(* IEC 61131-3 sources: stf-hw/stf-cad/line2/plc, 16 files *)

(* ---- DUT_PhysicalAI.st ---- *)
// timestamped I/O and the record every learned model is trained on
TYPE ST_TsInput : STRUCT bNewEdge : BOOL; nTimestamp : ULINT; END_STRUCT; END_TYPE     // EL1252 (DC ns)
TYPE ST_TsOutput : STRUCT bArm : BOOL; nFireAt : ULINT; END_STRUCT; END_TYPE          // EL2252 (DC ns)
// station states: named types (an enumeration declared inline in a VAR block is not portable)
TYPE T_ZoneArray : ARRAY[0..2] OF LREAL; END_TYPE   // per oven zone (one named type: FB_Band -> FB_Oven)
TYPE E_PickState : (WAIT, TRACK, GRIP, LIFT, PLACE, RELEASE, HOME); END_TYPE
TYPE E_AirlockOut : (IDLE, CARRY_OUT, INNER_CLOSE, OUTER_OPEN, SWAP, OUTER_CLOSE, INNER_OPEN, CARRY_IN); END_TYPE
// the stations (DT-4b)
TYPE ST_DeltaJob : STRUCT              // PLC -> a delta's motion program: a new nJob starts the job
    nJob : INT; nPuck : INT; nCol : INT; nLane : INT;   // C: the band row (fRowPos) + column -> puck; A/B: puck -> lane
    fRowPos : LREAL; fStart : LREAL;                    // band mm of the row's cut; master mm to start at
END_STRUCT; END_TYPE
TYPE ST_QcResult : STRUCT nSeq : INT; nPuck : INT; nVerdict : INT; END_STRUCT; END_TYPE   // edge PC: 1 pass, 2 reject
TYPE ST_Puck : STRUCT
    bFull : BOOL; bKicked : BOOL; bPending : BOOL;      // pending: a pick is decided, its grip not yet known
    nFlav : INT; nCol : INT; nVerdict : INT; fRowPos : LREAL;
END_STRUCT; END_TYPE
TYPE T_PuckArray : ARRAY[0..47] OF ST_Puck; END_TYPE
TYPE ST_Lane : STRUCT fBlock : LREAL; fPackAt : LREAL; nPackReq : INT; bCanPack : BOOL; END_STRUCT; END_TYPE   // s (master)
TYPE T_LaneArray : ARRAY[0..2] OF ST_Lane; END_TYPE
TYPE ST_PuckEvent : STRUCT
    nPuck : UINT; sNfc : STRING(16); nDcTime : ULINT; fMasterPos : LREAL;
    eStation : E_Station; aSignals : ARRAY[0..15] OF REAL; nImageId : UDINT; eOutcome : E_Outcome;
END_STRUCT; END_TYPE

(* ---- GVL_IO.st ---- *)
// GVL_IO - generated by plc_io.py from line_model: every signal, mapped in the I/O tree
{attribute 'qualified_only'}
VAR_GLOBAL
    axQ1                            : AXIS_REF;   // -KF20 ch1      M1_master_drive              stepper 17HS19-2004D-E1000+PG27
    encB1                    AT %I* : UDINT;   // -KF18 ch1      B1_master_encoder            master encoder, 1024 ppr RS422
    axQ41                           : AXIS_REF;   // -KF21 ch1      M_dep_rolls                  stepper 17HS19-2004D-E1000+PG27
    iolIOL1                  AT %I* : INT;   // -KF14 ch1      dep_hopper_level             ToF level (IO-Link)
    qQ2                      AT %Q* : BOOL;   // -KF5 ch7       top_cyl_weiss                valve coil (ISO6432-16x25)
    iQ2_S1                   AT %I* : BOOL;   // -KF1 ch1       top_cyl_weiss                reed switch retracted (ISO6432-16x25)
    iQ2_S2                   AT %I* : BOOL;   // -KF1 ch2       top_cyl_weiss                reed switch extended (ISO6432-16x25)
    qQ3                      AT %Q* : BOOL;   // -KF5 ch8       top_cyl_rot                  valve coil (ISO6432-16x25)
    iQ3_S1                   AT %I* : BOOL;   // -KF1 ch3       top_cyl_rot                  reed switch retracted (ISO6432-16x25)
    iQ3_S2                   AT %I* : BOOL;   // -KF1 ch4       top_cyl_rot                  reed switch extended (ISO6432-16x25)
    qQ4                      AT %Q* : BOOL;   // -KF5 ch9       top_cyl_blau                 valve coil (ISO6432-16x25)
    iQ4_S1                   AT %I* : BOOL;   // -KF1 ch5       top_cyl_blau                 reed switch retracted (ISO6432-16x25)
    iQ4_S2                   AT %I* : BOOL;   // -KF1 ch6       top_cyl_blau                 reed switch extended (ISO6432-16x25)
    iolIOL5                  AT %I* : INT;   // -KF14 ch2      top_level_weiss              ToF level (IO-Link)
    iolIOL6                  AT %I* : INT;   // -KF14 ch3      top_level_rot                ToF level (IO-Link)
    iolIOL7                  AT %I* : INT;   // -KF14 ch4      top_level_blau               ToF level (IO-Link)
    axQ40                           : AXIS_REF;   // -KF22 ch1      M_band                       stepper 17HS19-2004D-E1000+PG27
    qE1T1                    AT %Q* : BOOL;   // -KF5 ch12      oven_heater_E1T1             oven element SSR (500 W 230 V, L1)
    qE1T2                    AT %Q* : BOOL;   // -KF5 ch13      oven_heater_E1T2             oven element SSR (500 W 230 V, L2)
    qE1T3                    AT %Q* : BOOL;   // -KF5 ch14      oven_heater_E1T3             oven element SSR (500 W 230 V, L3)
    qE1B1                    AT %Q* : BOOL;   // -KF5 ch10      oven_heater_E1B1             oven element SSR (500 W 230 V, L1)
    qE1B2                    AT %Q* : BOOL;   // -KF5 ch11      oven_heater_E1B2             oven element SSR (500 W 230 V, L2)
    qQF1                     AT %Q* : BOOL;   // -KF6 ch7       oven_fan_1_motor             oven circulation fan 230 V 35 W (L2), coupling relay
    tcTC1                    AT %I* : INT;   // -KF12 ch1      oven_tc_1                    oven zone thermocouple K (duplex: this element -> PID)
    qE2T1                    AT %Q* : BOOL;   // -KF5 ch16      oven_heater_E2T1             oven element SSR (500 W 230 V, L3)
    qE2B1                    AT %Q* : BOOL;   // -KF5 ch15      oven_heater_E2B1             oven element SSR (350 W 230 V, L2)
    qQF2                     AT %Q* : BOOL;   // -KF6 ch8       oven_fan_2_motor             oven circulation fan 230 V 35 W (L3), coupling relay
    tcTC2                    AT %I* : INT;   // -KF12 ch2      oven_tc_2                    oven zone thermocouple K (duplex: this element -> PID)
    qE3T1                    AT %Q* : BOOL;   // -KF6 ch2       oven_heater_E3T1             oven element SSR (500 W 230 V, L1)
    qE3B1                    AT %Q* : BOOL;   // -KF6 ch1       oven_heater_E3B1             oven element SSR (350 W 230 V, L3)
    qQF3                     AT %Q* : BOOL;   // -KF6 ch9       oven_fan_3_motor             oven circulation fan 230 V 35 W (L2), coupling relay
    tcTC3                    AT %I* : INT;   // -KF12 ch3      oven_tc_3                    oven zone thermocouple K (duplex: this element -> PID)
    qQX1                     AT %Q* : BOOL;   // -KF6 ch10      oven_exhaust_fan             oven vapour exhaust fan 24 V EC
    aiIR1                    AT %I* : INT;   // -KF9 ch4       IR1_pyrometer                product temperature 0..10 V
    qQC1                     AT %Q* : BOOL;   // -KF6 ch3       cool_fan_1                   band cooling fan 24 V
    qQC2                     AT %Q* : BOOL;   // -KF6 ch4       cool_fan_2                   band cooling fan 24 V
    qQC3                     AT %Q* : BOOL;   // -KF6 ch5       cool_exfan_1                 band cooling fan 24 V
    qQC4                     AT %Q* : BOOL;   // -KF6 ch6       cool_exfan_2                 band cooling fan 24 V
    axdelta_C_M60                   : AXIS_REF;   // -KF25 ch1      delta_C_motor_60             stepper 17HS19-2004D-E1000+SWG17-30
    axdelta_C_M180                  : AXIS_REF;   // -KF23 ch1      delta_C_motor_180            stepper 17HS19-2004D-E1000+SWG17-30
    axdelta_C_M300                  : AXIS_REF;   // -KF24 ch1      delta_C_motor_300            stepper 17HS19-2004D-E1000+SWG17-30
    qdelta_C_VAC             AT %Q* : BOOL;   // -KF6 ch11      delta_C_cup_a                vacuum ejector valve
    ioldelta_C_VAC_P         AT %I* : INT;   // -KF15 ch2      delta_C_cup_a                vacuum level (analogue grip quality)
    iI1                      AT %I* : BOOL;   // -KF1 ch13      I1_full_check                puck already full (recirculating) -> delta C does NOT place
    iolNFC_W                 AT %I* : ARRAY[0..31] OF BYTE;   // -KF15 ch1      nfc_writer                   RFID/NFC head (IO-Link)
    itsI9                    AT %I* : ST_TsInput;   // -KF43 ch1      I9_landing_check             landing check after the place: is the cookie seated in the n
    qtsCAM1_TRG              AT %Q* : ST_TsOutput;   // -KF44 ch1      qc_camera                    camera trigger (timestamped)
    qQ17                     AT %Q* : BOOL;   // -KF6 ch12      qc_ringlight                 ring light 24 V
    aiAI1_R                  AT %I* : INT;   // -KF10 ch3      A1_colour_sensor             colour R 0..10 V
    aiAI1_G                  AT %I* : INT;   // -KF10 ch2      A1_colour_sensor             colour G 0..10 V
    aiAI1_B                  AT %I* : INT;   // -KF10 ch1      A1_colour_sensor             colour B 0..10 V
    iolNFC_W2                AT %I* : ARRAY[0..31] OF BYTE;   // -KF15 ch4      nfc_qc                       RFID/NFC head (IO-Link)
    qQ18                     AT %Q* : BOOL;   // -KF6 ch13      kick_cylinder                valve coil (ISO6432-10x100)
    iQ18_S1                  AT %I* : BOOL;   // -KF1 ch14      kick_cylinder                reed switch retracted (ISO6432-10x100)
    iQ18_S2                  AT %I* : BOOL;   // -KF1 ch15      kick_cylinder                reed switch extended (ISO6432-10x100)
    iolIOL4                  AT %I* : INT;   // -KF15 ch3      reject_level                 ToF level (IO-Link)
    axdelta_A_M_15                  : AXIS_REF;   // -KF26 ch1      delta_A_motor_-15            stepper 17HS19-2004D-E1000+SWG17-30
    axdelta_A_M105                  : AXIS_REF;   // -KF27 ch1      delta_A_motor_105            stepper 17HS19-2004D-E1000+SWG17-30
    axdelta_A_M225                  : AXIS_REF;   // -KF28 ch1      delta_A_motor_225            stepper 17HS19-2004D-E1000+SWG17-30
    qdelta_A_VAC             AT %Q* : BOOL;   // -KF6 ch14      delta_A_cup_a                vacuum ejector valve
    ioldelta_A_VAC_P         AT %I* : INT;   // -KF16 ch2      delta_A_cup_a                vacuum level (analogue grip quality)
    axdelta_B_M165                  : AXIS_REF;   // -KF29 ch1      delta_B_motor_165            stepper 17HS19-2004D-E1000+SWG17-30
    axdelta_B_M285                  : AXIS_REF;   // -KF30 ch1      delta_B_motor_285            stepper 17HS19-2004D-E1000+SWG17-30
    axdelta_B_M405                  : AXIS_REF;   // -KF31 ch1      delta_B_motor_405            stepper 17HS19-2004D-E1000+SWG17-30
    qdelta_B_VAC             AT %Q* : BOOL;   // -KF6 ch15      delta_B_cup_a                vacuum ejector valve
    ioldelta_B_VAC_P         AT %I* : INT;   // -KF16 ch3      delta_B_cup_a                vacuum level (analogue grip quality)
    qtsCAM2_TRG              AT %Q* : ST_TsOutput;   // -KF44 ch2      track_camera                 camera trigger (timestamped)
    iolNFC_R                 AT %I* : ARRAY[0..31] OF BYTE;   // -KF16 ch1      nfc_pick                     RFID/NFC head (IO-Link)
    axQ20                           : AXIS_REF;   // -KF32 ch1      lane_weiss_frame             stepper mini belt conveyor 60, end drive 17HS19-2004D-E1000+PG5 inside the frame
    qQ33                     AT %Q* : BOOL;   // -KF7 ch3       boxmag_weiss_fork_l          valve coil (ISO6432-8x10)
    iQ33_S1                  AT %I* : BOOL;   // -KF3 ch2       boxmag_weiss_fork_l          reed switch retracted (ISO6432-8x10)
    iQ33_S2                  AT %I* : BOOL;   // -KF3 ch3       boxmag_weiss_fork_l          reed switch extended (ISO6432-8x10)
    qQ36                     AT %Q* : BOOL;   // -KF7 ch6       sealer_weiss_head            sealing head DC SSR (24 V 60 W)
    tcQ36_TC                 AT %I* : INT;   // -KF12 ch4      sealer_weiss_head            sealing head thermocouple (integrated)
    axQ21                           : AXIS_REF;   // -KF33 ch1      lane_rot_frame               stepper mini belt conveyor 60, end drive 17HS19-2004D-E1000+PG5 inside the frame
    qQ34                     AT %Q* : BOOL;   // -KF7 ch4       boxmag_rot_fork_l            valve coil (ISO6432-8x10)
    iQ34_S1                  AT %I* : BOOL;   // -KF3 ch4       boxmag_rot_fork_l            reed switch retracted (ISO6432-8x10)
    iQ34_S2                  AT %I* : BOOL;   // -KF3 ch5       boxmag_rot_fork_l            reed switch extended (ISO6432-8x10)
    qQ37                     AT %Q* : BOOL;   // -KF7 ch7       sealer_rot_head              sealing head DC SSR (24 V 60 W)
    tcQ37_TC                 AT %I* : INT;   // -KF13 ch1      sealer_rot_head              sealing head thermocouple (integrated)
    axQ22                           : AXIS_REF;   // -KF34 ch1      lane_blau_frame              stepper mini belt conveyor 60, end drive 17HS19-2004D-E1000+PG5 inside the frame
    qQ35                     AT %Q* : BOOL;   // -KF7 ch5       boxmag_blau_fork_l           valve coil (ISO6432-8x10)
    iQ35_S1                  AT %I* : BOOL;   // -KF3 ch6       boxmag_blau_fork_l           reed switch retracted (ISO6432-8x10)
    iQ35_S2                  AT %I* : BOOL;   // -KF3 ch7       boxmag_blau_fork_l           reed switch extended (ISO6432-8x10)
    qQ38                     AT %Q* : BOOL;   // -KF7 ch8       sealer_blau_head             sealing head DC SSR (24 V 60 W)
    tcQ38_TC                 AT %I* : INT;   // -KF13 ch2      sealer_blau_head             sealing head thermocouple (integrated)
    qQ24                     AT %Q* : BOOL;   // -KF6 ch16      stacker_lift_weiss           valve coil (ISO6432-16x30)
    iQ24_S1                  AT %I* : BOOL;   // -KF2 ch12      stacker_lift_weiss           reed switch retracted (ISO6432-16x30)
    iQ24_S2                  AT %I* : BOOL;   // -KF2 ch13      stacker_lift_weiss           reed switch extended (ISO6432-16x30)
    iI12                     AT %I* : BOOL;   // -KF2 ch9       stack_count_weiss            reed switch on the lift cylinder: lifts are counted, the cas
    qQ25                     AT %Q* : BOOL;   // -KF7 ch1       stacker_lift_rot             valve coil (ISO6432-16x30)
    iQ25_S1                  AT %I* : BOOL;   // -KF2 ch14      stacker_lift_rot             reed switch retracted (ISO6432-16x30)
    iQ25_S2                  AT %I* : BOOL;   // -KF2 ch15      stacker_lift_rot             reed switch extended (ISO6432-16x30)
    iI13                     AT %I* : BOOL;   // -KF2 ch10      stack_count_rot              reed switch on the lift cylinder: lifts are counted, the cas
    qQ26                     AT %Q* : BOOL;   // -KF7 ch2       stacker_lift_blau            valve coil (ISO6432-16x30)
    iQ26_S1                  AT %I* : BOOL;   // -KF2 ch16      stacker_lift_blau            reed switch retracted (ISO6432-16x30)
    iQ26_S2                  AT %I* : BOOL;   // -KF3 ch1       stacker_lift_blau            reed switch extended (ISO6432-16x30)
    iI14                     AT %I* : BOOL;   // -KF2 ch11      stack_count_blau             reed switch on the lift cylinder: lifts are counted, the cas
    axQ27                           : AXIS_REF;   // -KF35 ch1      M_shuttle_weiss              stepper 17HS19-2004D-E1000
    axQ28                           : AXIS_REF;   // -KF36 ch1      M_shuttle_rot                stepper 17HS19-2004D-E1000
    axQ29                           : AXIS_REF;   // -KF37 ch1      M_shuttle_blau               stepper 17HS19-2004D-E1000
    // SO Q19            -KF58 ch4      frl                          soft-start / dump valve: safe exhaust of all air (SF3)  [TwinSAFE]
    // SI Q19.FB         -KF53 ch3      frl                          dump valve position switch (exhausted)  [TwinSAFE]
    qtsCAM4_TRG              AT %Q* : ST_TsOutput;   // -KF45 ch1      CAM4_pack                    camera trigger (timestamped)
    iB10                     AT %I* : BOOL;   // -KF2 ch6       M_shuttle_weiss              shuttle weiss home  [implied, not in CAD]
    iB11                     AT %I* : BOOL;   // -KF2 ch7       M_shuttle_rot                shuttle rot home  [implied, not in CAD]
    iB12                     AT %I* : BOOL;   // -KF2 ch8       M_shuttle_blau               shuttle blau home  [implied, not in CAD]
    iB20                     AT %I* : BOOL;   // -KF1 ch10      delta_C_motor_60             delta_C_motor_60 arm index  [implied, not in CAD]
    iB21                     AT %I* : BOOL;   // -KF1 ch11      delta_C_motor_180            delta_C_motor_180 arm index  [implied, not in CAD]
    iB22                     AT %I* : BOOL;   // -KF1 ch12      delta_C_motor_300            delta_C_motor_300 arm index  [implied, not in CAD]
    iB23                     AT %I* : BOOL;   // -KF1 ch16      delta_A_motor_-15            delta_A_motor_-15 arm index  [implied, not in CAD]
    iB24                     AT %I* : BOOL;   // -KF2 ch1       delta_A_motor_105            delta_A_motor_105 arm index  [implied, not in CAD]
    iB25                     AT %I* : BOOL;   // -KF2 ch2       delta_A_motor_225            delta_A_motor_225 arm index  [implied, not in CAD]
    iB26                     AT %I* : BOOL;   // -KF2 ch3       delta_B_motor_165            delta_B_motor_165 arm index  [implied, not in CAD]
    iB27                     AT %I* : BOOL;   // -KF2 ch4       delta_B_motor_285            delta_B_motor_285 arm index  [implied, not in CAD]
    iB28                     AT %I* : BOOL;   // -KF2 ch5       delta_B_motor_405            delta_B_motor_405 arm index  [implied, not in CAD]
    aiBC1                    AT %I* : INT;   // -KF9 ch1                                    oven element feed L1 current 0..20 A (heater break)  [implied, not in CAD]
    aiBC2                    AT %I* : INT;   // -KF9 ch2                                    oven element feed L2 current 0..20 A (heater break)  [implied, not in CAD]
    aiBC3                    AT %I* : INT;   // -KF9 ch3                                    oven element feed L3 current 0..20 A (heater break)  [implied, not in CAD]
    // SI S20.A          -KF49 ch2      lock_S20                     door closed AND locked, OSSD A (SF2)  [TwinSAFE]
    // SI S20.B          -KF49 ch3      lock_S20                     door closed AND locked, OSSD B (SF2)  [TwinSAFE]
    // SO S20.UNL        -KF56 ch1      lock_S20                     unlock solenoid (power-to-unlock, only at standstill)  [TwinSAFE]
    // SI S21.A          -KF49 ch4      lock_S21                     door closed AND locked, OSSD A (SF2)  [TwinSAFE]
    // SI S21.B          -KF50 ch1      lock_S21                     door closed AND locked, OSSD B (SF2)  [TwinSAFE]
    // SO S21.UNL        -KF56 ch2      lock_S21                     unlock solenoid (power-to-unlock, only at standstill)  [TwinSAFE]
    // SI S22.A          -KF50 ch2      lock_S22                     door closed AND locked, OSSD A (SF2)  [TwinSAFE]
    // SI S22.B          -KF50 ch3      lock_S22                     door closed AND locked, OSSD B (SF2)  [TwinSAFE]
    // SO S22.UNL        -KF56 ch3      lock_S22                     unlock solenoid (power-to-unlock, only at standstill)  [TwinSAFE]
    // SI Q42.CLA        -KF46 ch1      trapdoor_weiss               trapdoor closed, safety sensor OSSD A  [TwinSAFE]
    // SI Q42.CLB        -KF46 ch2      trapdoor_weiss               trapdoor closed, safety sensor OSSD B  [TwinSAFE]
    qQ42                     AT %Q* : BOOL;   // -KF5 ch1       trapdoor_weiss               trapdoor valve (spring-return closes on exhaust)
    // SI Q43.CLA        -KF46 ch3      trapdoor_rot                 trapdoor closed, safety sensor OSSD A  [TwinSAFE]
    // SI Q43.CLB        -KF46 ch4      trapdoor_rot                 trapdoor closed, safety sensor OSSD B  [TwinSAFE]
    qQ43                     AT %Q* : BOOL;   // -KF5 ch2       trapdoor_rot                 trapdoor valve (spring-return closes on exhaust)
    // SI Q44.CLA        -KF47 ch1      trapdoor_blau                trapdoor closed, safety sensor OSSD A  [TwinSAFE]
    // SI Q44.CLB        -KF47 ch2      trapdoor_blau                trapdoor closed, safety sensor OSSD B  [TwinSAFE]
    qQ44                     AT %Q* : BOOL;   // -KF5 ch3       trapdoor_blau                trapdoor valve (spring-return closes on exhaust)
    // SI S30.A          -KF50 ch4      aldoor_boxes                 boxes airlock outer door closed AND locked, OSSD A  [TwinSAFE]
    // SI S30.B          -KF51 ch1      aldoor_boxes                 boxes airlock outer door closed AND locked, OSSD B  [TwinSAFE]
    // SO S30.UNL        -KF56 ch4      aldoor_boxes                 boxes airlock outer door lock release (interlocked)  [TwinSAFE]
    qS30_DRV                 AT %Q* : BOOL;   // -KF5 ch4       aldoor_boxes                 boxes airlock outer door drive valve (force-limited)
    // SI S32.A          -KF51 ch4      aldoor_inner                 out airlock inner door closed AND locked, OSSD A  [TwinSAFE]
    // SI S32.B          -KF52 ch1      aldoor_inner                 out airlock inner door closed AND locked, OSSD B  [TwinSAFE]
    // SO S32.UNL        -KF57 ch2      aldoor_inner                 out airlock inner door lock release (interlocked)  [TwinSAFE]
    qS32_DRV                 AT %Q* : BOOL;   // -KF5 ch6       aldoor_inner                 out airlock inner door drive valve (force-limited)
    // SI S31.A          -KF51 ch2      aldoor_out                   out airlock outer door closed AND locked, OSSD A  [TwinSAFE]
    // SI S31.B          -KF51 ch3      aldoor_out                   out airlock outer door closed AND locked, OSSD B  [TwinSAFE]
    // SO S31.UNL        -KF57 ch1      aldoor_out                   out airlock outer door lock release (interlocked)  [TwinSAFE]
    qS31_DRV                 AT %Q* : BOOL;   // -KF5 ch5       aldoor_out                   out airlock outer door drive valve (force-limited)
    // SI S10.A          -KF47 ch3      estop_S10_head               E-stop NC contact A (SF1, 2-channel)  [TwinSAFE]
    // SI S10.B          -KF47 ch4      estop_S10_head               E-stop NC contact B (SF1, 2-channel)  [TwinSAFE]
    // SI S11.A          -KF48 ch1      estop_S11_head               E-stop NC contact A (SF1, 2-channel)  [TwinSAFE]
    // SI S11.B          -KF48 ch2      estop_S11_head               E-stop NC contact B (SF1, 2-channel)  [TwinSAFE]
    // SI S12.A          -KF48 ch3      estop_S12_head               E-stop NC contact A (SF1, 2-channel)  [TwinSAFE]
    // SI S12.B          -KF48 ch4      estop_S12_head               E-stop NC contact B (SF1, 2-channel)  [TwinSAFE]
    // SI S13            -KF49 ch1      reset_S13_head               reset pushbutton (manual reset on the falling edge)  [TwinSAFE]
    iBOXES_DOCK1             AT %I* : BOOL;   // -KF3 ch11      port_boxes                   AMR docked at boxes (1)  [implied, not in CAD]
    iBOXES_DOCK2             AT %I* : BOOL;   // -KF3 ch12      port_boxes                   AMR docked at boxes (2)  [implied, not in CAD]
    iOUT_DOCK1               AT %I* : BOOL;   // -KF3 ch13      port_out                     AMR docked at out (1)  [implied, not in CAD]
    iOUT_DOCK2               AT %I* : BOOL;   // -KF3 ch14      port_out                     AMR docked at out (2)  [implied, not in CAD]
    // SI S34.A          -KF52 ch2      reject_bin_wall_front        reject drawer in place, OSSD A  [TwinSAFE]
    // SI S34.B          -KF52 ch3      reject_bin_wall_front        reject drawer in place, OSSD B  [TwinSAFE]
    // SO K1             -KF57 ch3                                   contactor coil: 48 V motor supply, channel 1 (all EL7047)  [TwinSAFE]
    // SO K2             -KF57 ch4                                   contactor coil: 48 V motor supply, channel 2 (in series with K1)  [TwinSAFE]
    // SO K3             -KF58 ch1                                   contactor coil: 400 V oven feed + 24 V heater PSU, channel 1 (3-pole)  [TwinSAFE]
    // SO K4             -KF58 ch2                                   contactor coil: 400 V oven feed + 24 V heater PSU, channel 2 (in series with K3)  [TwinSAFE]
    // SO K5             -KF58 ch3                                   contactor coil: 48 V branch of the out-port zone (Q27, Q28, Q29)  [TwinSAFE]
    // SI K1K2.EDM       -KF52 ch4                                   EDM: K1 + K2 mirror contacts in series (welded contact detection)  [TwinSAFE]
    // SI K3K4.EDM       -KF53 ch1                                   EDM: K3 + K4 mirror contacts (welded contact detection)  [TwinSAFE]
    // SI K5.EDM         -KF53 ch2                                   EDM: K5 mirror contact (welded contact detection)  [TwinSAFE]
    // SO Y1             -KF59 ch1      valve_island                 safe exhaust of the boxes-port pressure zone (SF6)  [TwinSAFE]
    // SI Y1.FB          -KF53 ch4      valve_island                 boxes zone valve position switch (exhausted)  [TwinSAFE]
    iTC1_STL                 AT %I* : BOOL;   // -KF1 ch7       oven_tc_1                    safety temperature limiter tripped (SF4, own element of a duplex thermocouple; its contact is in the coil of zone contactor KH1)
    iTC2_STL                 AT %I* : BOOL;   // -KF1 ch8       oven_tc_2                    safety temperature limiter tripped (SF4, own element of a duplex thermocouple; its contact is in the coil of zone contactor KH2)
    iTC3_STL                 AT %I* : BOOL;   // -KF1 ch9       oven_tc_3                    safety temperature limiter tripped (SF4, own element of a duplex thermocouple; its contact is in the coil of zone contactor KH3)
    iQ36_STL                 AT %I* : BOOL;   // -KF3 ch8       sealer_weiss_head            safety temperature limiter tripped (SF4, own element of a duplex thermocouple; its relay contact is in the heater load path)
    iQ37_STL                 AT %I* : BOOL;   // -KF3 ch9       sealer_rot_head              safety temperature limiter tripped (SF4, own element of a duplex thermocouple; its relay contact is in the heater load path)
    iQ38_STL                 AT %I* : BOOL;   // -KF3 ch10      sealer_blau_head             safety temperature limiter tripped (SF4, own element of a duplex thermocouple; its relay contact is in the heater load path)
    axMasterEnc                     : AXIS_REF;   // NC encoder axis on B1: the virtual master (gearing, cams)
    xSafeRunPermit           AT %I* : BOOL;   // EL6910 standard process data: no stop demand, doors locked, resets done
    stDeltaC                        : ST_DeltaJob;   // delta C: the job its motion program (kinematic group + conveyor tracking) executes
    stDeltaA                        : ST_DeltaJob;   // delta A: the job its motion program (kinematic group + conveyor tracking) executes
    stDeltaB                        : ST_DeltaJob;   // delta B: the job its motion program (kinematic group + conveyor tracking) executes
    stQc                            : ST_QcResult;   // the QC verdict, written by the edge PC (ADS) per puck
    xHmiLoad                 AT %I* : BOOL;   // HMI start of production: load cookies into the pucks
END_VAR

(* ---- F_InSlice.st ---- *)
// F_InSlice - TRUE while fPhase (0..1 of the PWM period) lies in [fStart, fStart + fDuty), wrapping at 1
FUNCTION F_InSlice : BOOL
VAR_INPUT fPhase, fStart, fDuty : LREAL; END_VAR
F_InSlice := LMOD(fPhase - fStart + 1.0, 1.0) < fDuty;

(* ---- FB_Airlock.st ---- *)
// FB_Airlock - standard-side sequence of the two AMR airlocks. It only REQUESTS; the TwinSAFE
// project (SF6) refuses any unlock that breaks the interlock, so a bug here cannot open both sides.
//
// OUT (cassettes), per lane, started by the lift counter 75 s before full (the AMR is called then):
//   1 carrier: full cassette stacker -> chamber (200 mm at 100 mm/s)
//   2 request S32 close + lock (inner door); TwinSAFE drops K5 (shuttles)
//   3 AMR docked (OUT.DOCK1/2) -> request S31 unlock + open (outer door)
//   4 AMR swaps full <-> empty (20 s [assumed]); S31 close + lock
//   5 request S32 unlock + open; K5 on; carrier: empty chamber -> stacker
//   exchange 30 s; the stacker platform holds 1 sealed pack meanwhile, so a robot on
//   time costs no production. Lanes run a third of a fill apart (CASS_STAGGER) so exchanges never coincide.
// BOXES (tray stacks): AMR docked -> trapdoors closed (Q42..Q44.CL) + Y1 exhausted -> S30 unlock + open;
//   AMR sets stacks in the chamber; S30 close + lock -> Y1 on -> trapdoor over each low magazine drops its stack.
FUNCTION_BLOCK FB_Airlock
VAR_INPUT nLaneFull : INT; bAmrDocked : BOOL; END_VAR
VAR eOut : E_AirlockOut; END_VAR

(* ---- FB_Arrivals.st ---- *)
// FB_Arrivals - the pucks passing ONE station of the loop, from the master position alone: puck k is at the
// station when the master is at fStation - k x 80 (mod 3840.037061436, the loop); after puck k comes puck k-1.
// The arrival is reported in the scan the master passes it, with the EXACT position it happened at (fArr).
FUNCTION_BLOCK FB_Arrivals
VAR_INPUT fMaster : LREAL; fStation : LREAL; END_VAR
VAR_OUTPUT bArrive : BOOL; nPuck : INT; fArr : LREAL; END_VAR
VAR bInit : BOOL; nNext, k : INT; fNext, f : LREAL; END_VAR
bArrive := FALSE;
IF NOT bInit THEN                          // the first arrival from now on, over all 48 pucks
    fNext := fMaster + 3840.037061436;
    FOR k := 0 TO 47 DO
        f := fMaster + LMOD(fStation - INT_TO_LREAL(k) * 80.0 - fMaster, 3840.037061436);
        IF f < fNext THEN fNext := f;  nNext := k; END_IF;
    END_FOR;
    bInit := TRUE;
END_IF;
IF fMaster >= fNext THEN
    bArrive := TRUE;  nPuck := nNext;  fArr := fNext;
    nNext := (nNext + 47) MOD 48;
    fNext := fArr + LMOD(fStation - INT_TO_LREAL(nNext) * 80.0 - fArr, 3840.037061436);
END_IF;

(* ---- FB_Band.st ---- *)
// FB_Band - the mesh band (2.292 mm/s) and the depositor rolls are GEARED to the master axis:
// one row of 6 per 6 pucks (24 s). The wire is cammed from the rolls.
// Topping: rows k and k+3 get flavour k (Q2/Q3/Q4), 100 mm after the die.
// A cold oven (bOvenReady FALSE) stops the depositor, never the band: what is in the oven bakes out.
// aZoneContent (the oven's feed-forward): every row the depositor cuts (the rolls' measured motion, AND dough in the
// hopper - IOL1) is remembered at the band position of its cut; a zone's content = the rows between its walls / the
// 3.69 rows a full zone holds. Turning rolls on an empty hopper cut nothing (DT-4a finding 15).
FUNCTION_BLOCK FB_Band
VAR_IN_OUT axBand : AXIS_REF; axRolls : AXIS_REF; axMaster : AXIS_REF; END_VAR   // by reference (MC blocks)
VAR_INPUT bOvenReady : BOOL; nDoughLevel : INT; END_VAR   // nDoughLevel: IOL1 distance to the dough, 0.1 mm
VAR_OUTPUT fPos : LREAL; aZoneContent : T_ZoneArray;   // 0..1 per zone, from the rows cut
    nRows : UDINT; fRowPos : LREAL;        // rows cut so far, the band position of the last (-> FB_Transfer)
END_VAR
VAR RETAIN                                 // the rows on the band survive a power cycle (they are still there)
    aCut : ARRAY[0..31] OF LREAL;          // band position of each row cut (ring), -1 = empty
    nCut : INT; fLastCut : LREAL; bFirst : BOOL := TRUE;
END_VAR
VAR fbGearBand, fbGearRolls : MC_GearIn; fbGearOutRolls : MC_GearOut; fbHaltRolls : MC_Halt;
    k, i : INT; d : LREAL; fDough : LREAL;   // kg of dough in the hopper
    fDoughRow : LREAL;                     // the most dough seen while this row was pressed out
    aZoneOff : ARRAY[0..2] OF LREAL := [200.0, 403.0, 606.0];   // die -> zone start, mm of band
END_VAR
fbGearBand(Master := axMaster, Slave := axBand, Execute := TRUE, RatioNumerator := 2.291666666667,
           RatioDenominator := 20);   // band mm/s per master mm/s: exact (rounded, rows drift: finding 17)
fbGearRolls(Master := axMaster, Slave := axRolls, Execute := bOvenReady, RatioNumerator := 1.0, RatioDenominator := 1);
// a FALLING Execute does not decouple a geared slave (PLCopen): oven not ready -> decouple the rolls, then brake them
fbGearOutRolls(Slave := axRolls, Execute := NOT bOvenReady);
fbHaltRolls(Axis := axRolls, Execute := NOT bOvenReady AND fbGearOutRolls.Done, Deceleration := 40.0);
fPos := axBand.NcToPlc.ActPos;
fDough := (276.0 - INT_TO_LREAL(nDoughLevel) * 0.1) * 0.111090;
fDoughRow := MAX(fDoughRow, fDough);       // the level drops as the slug leaves: judge the row on the level before
IF bFirst THEN
    FOR i := 0 TO 31 DO aCut[i] := -1.0; END_FOR;
    fLastCut := fPos;  bFirst := FALSE;
END_IF;
IF fPos - fLastCut >= 55.0000 THEN                  // one row pitch of band: the wire cuts a row if the rolls run
    fLastCut := fLastCut + 55.0000;
    // a row exists if the rolls REALLY turned (their actual velocity), not if they were told to: a halt brakes;
    // and only from a hopper holding a row's dough (6 x 0.0112 kg)
    IF ABS(axRolls.NcToPlc.ActVelo) > 0.0 AND fDoughRow >= 0.0672 THEN
        aCut[nCut] := fLastCut;  nCut := (nCut + 1) MOD 32;  nRows := nRows + 1;  fRowPos := fLastCut;
    END_IF;
    fDoughRow := fDough;
END_IF;
FOR k := 0 TO 2 DO
    aZoneContent[k] := 0.0;
    FOR i := 0 TO 31 DO
        IF aCut[i] >= 0.0 THEN
            d := fPos - aCut[i];
            IF d >= aZoneOff[k] AND d < aZoneOff[k] + 203.0 THEN
                aZoneContent[k] := aZoneContent[k] + 0.270936;
            END_IF;
        END_IF;
    END_FOR;
    aZoneContent[k] := MIN(aZoneContent[k], 1.0);
END_FOR;

(* ---- FB_CameraTrigger.st ---- *)
// FB_CameraTrigger - fire every camera at a puck's master position via EL2252 (DC time), so each image
// is exactly aligned with the puck (NFC id), the master position and every other sensor sample.
FUNCTION_BLOCK FB_CameraTrigger
VAR_INPUT fMasterPos : LREAL; fTriggerPos : LREAL; END_VAR
VAR_IN_OUT stOut : ST_TsOutput; END_VAR
// nFireAt := DC time now + (fTriggerPos - fMasterPos) / 20 mm/s -> the terminal fires on the ns

(* ---- FB_DeltaPicker.st ---- *)
// FB_DeltaPicker - conveyor tracking pick of a moving cookie, place into the lane pocket.
// Kinematics: the NC delta transformation (TF5110-class, licence to confirm) with conveyor tracking coupled to the
// master axis executes stJob (the puck, the lane, the master position to start at). A is upstream and picks; B
// catches what A missed (N+1). Placement budget: backlash + steps <= DELTA_REP (line_model.sizing, the Jacobian).
// A passing pass-verdict cookie is taken if the delta is free (after its last pick, 2 s) and its lane is not
// indexing, early enough to grip (0.8 s) before the puck leaves the reach; else B counts it missed (it
// recirculates). The grip is known from the vacuum at T_GRAB: the pick is booked when it is decided (the tray fill,
// a full tray indexes the lane: blocked 2 s) and taken back if the cup holds nothing.
FUNCTION_BLOCK FB_DeltaPicker
VAR_IN_OUT stJob : ST_DeltaJob; aPuck : T_PuckArray; aLane : T_LaneArray; END_VAR
VAR_INPUT fMaster : LREAL; nDelta : INT; fIn : LREAL; fOut : LREAL; nVacuum : INT; END_VAR
VAR_OUTPUT bVacuum : BOOL; bMissed : BOOL; nPicks, nPickFail, nMissed, nRollback : DINT; END_VAR
VAR fbArr : FB_Arrivals; pk, f, q : INT; t, tOut, tStart, tNow, fBusy, fHold : LREAL;
    aFill : ARRAY[0..2] OF INT;            // cookies in this delta's tray, per lane
    aQPuck, aQLane : ARRAY[0..3] OF INT; aQStart, aQPrev : ARRAY[0..3] OF LREAL; aQPack : ARRAY[0..3] OF BOOL;
    nQHead, nQTail : INT;                  // the jobs given to the delta, not yet gripped
END_VAR
tNow := fMaster / 20.0;
fbArr(fMaster := fMaster, fStation := fIn);
bMissed := FALSE;
IF fbArr.bArrive THEN
    pk := fbArr.nPuck;
    IF aPuck[pk].bFull AND NOT aPuck[pk].bPending AND NOT aPuck[pk].bKicked AND aPuck[pk].nVerdict = 1 THEN
        f := aPuck[pk].nFlav;
        t := fbArr.fArr / 20.0;
        tOut := t + (fOut - fIn) / 20.0;
        tStart := MAX(t, MAX(fBusy, aLane[f].fBlock));
        IF tStart + 0.8 <= tOut AND aLane[f].bCanPack THEN
            fBusy := tStart + 2.0;
            stJob.nPuck := pk;  stJob.nCol := aPuck[pk].nCol;  stJob.nLane := f;  stJob.fRowPos := aPuck[pk].fRowPos;
            stJob.fStart := tStart * 20.0;  stJob.nJob := (stJob.nJob + 1) MOD 10000;
            aPuck[pk].bPending := TRUE;
            aQPuck[nQTail] := pk;  aQLane[nQTail] := f;  aQStart[nQTail] := tStart;  aQPack[nQTail] := FALSE;
            aFill[f] := aFill[f] + 1;
            IF aFill[f] >= 3 THEN       // the tray is full: the lane indexes when this pick ends
                aFill[f] := 0;  aQPack[nQTail] := TRUE;  aQPrev[nQTail] := aLane[f].fBlock;
                aLane[f].fBlock := fBusy + 2.0;  aLane[f].fPackAt := fBusy;
                aLane[f].nPackReq := aLane[f].nPackReq + 1;
            END_IF;
            nQTail := (nQTail + 1) MOD 4;
        ELSIF nDelta = 1 THEN
            bMissed := TRUE;  nMissed := nMissed + 1;
        END_IF;
    END_IF;
END_IF;
IF nQHead <> nQTail THEN                   // the grip of the oldest job
    IF tNow >= aQStart[nQHead] + 0.8 THEN
        pk := aQPuck[nQHead];  f := aQLane[nQHead];
        IF nVacuum <= -300 THEN
            aPuck[pk].bFull := FALSE;  aPuck[pk].bPending := FALSE;  nPicks := nPicks + 1;
            fHold := aQStart[nQHead] + 2.0;   // held until it is placed
        ELSE                               // not held: the cookie rides on, the booking is taken back
            aPuck[pk].bPending := FALSE;  nPickFail := nPickFail + 1;
            IF aQPack[nQHead] THEN
                aFill[f] := 2;  aLane[f].fBlock := aQPrev[nQHead];  aLane[f].nPackReq := aLane[f].nPackReq - 1;
            ELSE
                aFill[f] := aFill[f] - 1;
            END_IF;
            q := (nQHead + 1) MOD 4;       // a later job of this delta already booked on the taken-back fill
            IF q <> nQTail THEN nRollback := nRollback + 1; END_IF;
        END_IF;
        nQHead := (nQHead + 1) MOD 4;
    END_IF;
END_IF;
bVacuum := tNow < fHold;
IF nQHead <> nQTail THEN
    IF tNow >= aQStart[nQHead] THEN bVacuum := TRUE; END_IF;
END_IF;

(* ---- FB_Lane.st ---- *)
// FB_Lane - index one tray pitch (160 mm in 1.6 s) when a tray is full, as the pick that filled it ends;
// the pickers keep off the lane meanwhile (2 s). Seal in the index pause (1 s <= 2 s);
// stacker lifts each pack through the pawls; the lift counter says 'cassette full' at 27 packs;
// shuttle swap (OPEN DESIGN ISSUE: a single bar cannot exchange two cassettes - see joints/README).
// bCanPack: TRUE until the logistics (tray magazine, cassette, airlock) are written (DT-4b part 2).
FUNCTION_BLOCK FB_Lane
VAR_IN_OUT axLane : AXIS_REF; stLane : ST_Lane; END_VAR
VAR_INPUT fMaster : LREAL; END_VAR
VAR_OUTPUT nPacks : DINT; END_VAR
VAR fbPower : MC_Power; fbIndex : MC_MoveRelative; nDone : INT; bGo : BOOL; END_VAR
fbPower(Axis := axLane, Enable := TRUE, Enable_Positive := TRUE, Enable_Negative := FALSE);
stLane.bCanPack := TRUE;
bGo := stLane.nPackReq > nDone AND fMaster / 20.0 >= stLane.fPackAt AND fbPower.Status;
fbIndex(Axis := axLane, Execute := bGo, Distance := 160.0, Velocity := 200.0,
        Acceleration := 250.0, Deceleration := 250.0);
IF fbIndex.Done THEN nDone := nDone + 1;  nPacks := nPacks + 1; END_IF;

(* ---- FB_MasterAxis.st ---- *)
// FB_MasterAxis - the electronic line shaft. The chain NEVER stops (no stop path in the
// automatic mode, only losses). v = 20 mm/s, pitch = 80 mm -> takt 4.00 s.
// The master position is the MEASURING-WHEEL encoder B1 (EL5101), not the drive's own encoder,
// so sprocket slip shows as a drift between the two (health signal).
FUNCTION_BLOCK FB_MasterAxis
VAR_IN_OUT                        // axes BY REFERENCE: MC blocks on a copy would never move the real axis
    axDrive  : AXIS_REF;          // Q1 on EL7047 (closed loop)
    axMaster : AXIS_REF;          // NC encoder axis on B1 (virtual master for gearing / cams)
END_VAR
VAR_INPUT
    nEncoder : UDINT;             // B1 counts
END_VAR
VAR_OUTPUT
    fPos     : LREAL;             // mm along the loop, modulo the loop length
    fAbs     : LREAL;             // mm since power-up (the stations' time base: tau = fAbs / v)
    fDrift   : LREAL;             // drive encoder - B1, mm (slip monitor)
END_VAR
VAR
    fbPower : MC_Power; fbVel : MC_MoveVelocity;
END_VAR
fbPower(Axis := axDrive, Enable := TRUE, Enable_Positive := TRUE, Enable_Negative := FALSE);
fbVel(Axis := axDrive, Execute := fbPower.Status, Velocity := 20.0, Acceleration := 20.0, Deceleration := 20.0,
      Direction := MC_Positive_Direction);
fPos := LMOD(axMaster.NcToPlc.ActPos, 3840.037061436);   // the chain's loop, not N x P (finding 16)
fAbs := axMaster.NcToPlc.ActPos;
fDrift := axDrive.NcToPlc.ActPos - axMaster.NcToPlc.ActPos;

(* ---- FB_Oven.st ---- *)
// FB_Oven - 3 zones. Per zone: FEED-FORWARD of the band load (from the band content FB_Band tracks,
// row by row) + PI on the zone TC (SIMC-tuned on the oven_ctrl.py model) with conditional-integration
// anti-windup -> 2 s time-proportioning PWM on every element SSR of the zone. Cold start: set point ramp
// 10 K/min with the ramp power fed forward.
// LEARNING feed-forward (upgrade V-1): calm at the set point (+-0.5 K for 120 s) on an empty band the PI
// share moves into aW0 (base load error, W), on a full band into aA1 (product load factor), time constant
// 600 s; the integrator gives the same amount back. Both are PERSISTENT (oven_ctrl S6: +-20 % model error).
// HEATER BREAK: current transducers BC1, BC2, BC3 on L1-L3 of the element feed. The expected phase current
// (every element in its PWM slice + the fans) lagged by the transducer's 0.3 s; short by > half the
// smallest element of the phase for 0.2 s -> alarm; the elements in their slice through the short are
// the candidates, an element seen conducting while the phase reads right is cleared -> named (oven_ctrl S4).
// A named element leaves its zone's model (power, gain); if the rest cannot carry the full load, bReady drops
// and FB_Band stops the depositor. The STB (SF4) is hardware.
//   Z1 210 C: TC TC1 -> E1T1 500 W top L1, E1T2 500 W top L2, E1T3 500 W top L3, E1B1 500 W bot L1, E1B2 500 W bot L2; fan QF1
//   Z2 200 C: TC TC2 -> E2T1 500 W top L3, E2B1 350 W bot L2; fan QF2
//   Z3 185 C: TC TC3 -> E3T1 500 W top L1, E3B1 350 W bot L3; fan QF3
// Steady load at 900 cookies/h: Z1 1516 W, Z2 563 W, Z3 562 W.
// The recipe holds +-2 K (oven.py bake window); bReady = every zone inside it for 60 s.
FUNCTION_BLOCK FB_Oven
VAR_INPUT  bRunEnable : BOOL; aContent : T_ZoneArray; END_VAR   // aContent: 0..1 zone filled (FB_Band)
VAR_OUTPUT bReady : BOOL; aTemp : ARRAY[0..2] OF LREAL; aDuty : ARRAY[0..2] OF LREAL;
           aElementAlarm : ARRAY[0..2] OF BOOL; aBroken : ARRAY[0..8] OF BOOL; bHold : BOOL;
           fPower_W : LREAL; END_VAR
VAR PERSISTENT
    aW0 : ARRAY[0..2] OF LREAL;                                   // W, learned base-load error
    aA1 : ARRAY[0..2] OF LREAL := [1.0, 1.0, 1.0];   // learned product-load factor
END_VAR
VAR
    aSet  : ARRAY[0..2] OF LREAL := [210.0, 200.0, 185.0];      // degC (oven.py recipe)
    aKc   : ARRAY[0..2] OF LREAL := [0.0225, 0.0650, 0.0673];  // 1/K
    aTi   : ARRAY[0..2] OF LREAL := [150.0, 152.0, 148.0];  // s
    aP    : ARRAY[0..2] OF LREAL := [2500.0, 850.0, 850.0];        // W installed
    aC    : ARRAY[0..2] OF LREAL := [2109.0, 2109.0, 2109.0];        // J/K
    aLoadEmpty : ARRAY[0..2] OF LREAL := [538.0, 23.0, 264.0];   // W, empty band
    aLoadFull  : ARRAY[0..2] OF LREAL := [1516.0, 563.0, 562.0];   // W, full band
    aSp, aI, aLost, aCalm : ARRAY[0..2] OF LREAL;   // aSp := aTemp at power-up (the ramp starts where the zone is)
    fRamp : LREAL := 0.1667;    // K/s
    // elements, flattened in slice order: zone, slice i of n, phase 0..2 = L1..L3, W
    aElZone  : ARRAY[0..8] OF INT := [0, 0, 0, 0, 0, 1, 1, 2, 2];
    aElSlice : ARRAY[0..8] OF LREAL := [0.0, 0.2, 0.4, 0.6, 0.8, 0.0, 0.5, 0.0, 0.5];   // i / n
    aElPh    : ARRAY[0..8] OF INT := [0, 1, 2, 0, 1, 2, 1, 0, 2];
    aElW     : ARRAY[0..8] OF LREAL := [500.0, 500.0, 500.0, 500.0, 500.0, 500.0, 350.0, 500.0, 350.0];
    aOn, aCand : ARRAY[0..8] OF BOOL;
    aFanA : ARRAY[0..2] OF LREAL := [0.000, 0.304, 0.152];   // A, fans on the feed
    aThrA : ARRAY[0..2] OF LREAL := [1.087, 0.761, 0.761];   // A, half the smallest element
    aExp, aExpLag, aMeas, aShort : ARRAY[0..2] OF LREAL;
    aPhAlarm, aShortOn : ARRAY[0..2] OF BOOL;
    aOnT : ARRAY[0..8] OF LREAL;  aRecent, aTry, aOnLast : ARRAY[0..8] OF BOOL;
    aSince, aAlarmT, aProbeT, aProbeMax : ARRAY[0..2] OF LREAL;
    aNamedT : ARRAY[0..2] OF LREAL := [-1.0E9, -1.0E9, -1.0E9];   // s: when the phase last named an element
    aProbe : ARRAY[0..2] OF INT := [-1, -1, -1];
    fNow_s, fPhase, dW, fProd : LREAL;     // fNow_s: task time in s, advanced every 10 ms cycle
    tStable : TON; k, i, j, n, m : INT; e, uff, u : LREAL; bRamp, bAnyAlarm, bSame, bSettled, bInit : BOOL;
END_VAR
fNow_s := fNow_s + 0.01;                   // the task clock (10 ms cycle): PWM phase + heater-break timing
aTemp[0] := INT_TO_LREAL(GVL_IO.tcTC1) / 10.0;
aTemp[1] := INT_TO_LREAL(GVL_IO.tcTC2) / 10.0;
aTemp[2] := INT_TO_LREAL(GVL_IO.tcTC3) / 10.0;
aMeas[0] := INT_TO_LREAL(GVL_IO.aiBC1) / 32767.0 * 20.0;   // A, L1
aMeas[1] := INT_TO_LREAL(GVL_IO.aiBC2) / 32767.0 * 20.0;   // A, L2
aMeas[2] := INT_TO_LREAL(GVL_IO.aiBC3) / 32767.0 * 20.0;   // A, L3
IF NOT bInit THEN                          // power-up: the set-point ramp starts where each zone IS (a hot
    FOR k := 0 TO 2 DO aSp[k] := aTemp[k]; END_FOR;   // oven restarts at its set point, a cold one ramps)
    bInit := TRUE;
END_IF;
bAnyAlarm := aPhAlarm[0] OR aPhAlarm[1] OR aPhAlarm[2] OR aElementAlarm[0] OR aElementAlarm[1] OR aElementAlarm[2];   // learning frozen until repaired
FOR k := 0 TO 2 DO
    aSp[k] := MIN(aSet[k], aSp[k] + fRamp * 0.01);  bRamp := aSp[k] < aSet[k];        // 10 ms task
    e := aSp[k] - aTemp[k];
    fProd := aContent[k] * (aLoadFull[k] - aLoadEmpty[k]);
    uff := (aLoadEmpty[k] + aW0[k] + aA1[k] * fProd + SEL(bRamp, 0.0, aC[k] * fRamp)) / (aP[k] - aLost[k]);
    u := uff + aKc[k] * aP[k] / (aP[k] - aLost[k]) * (e + aI[k] / aTi[k]);
    IF (u > 0.0 AND u < 1.0) OR (u >= 1.0 AND e < 0.0) OR (u <= 0.0 AND e > 0.0) THEN aI[k] := aI[k] + e * 0.01; END_IF;
    aDuty[k] := LIMIT(0.0, u, 1.0);
    // learning feed-forward
    IF ABS(e) < 0.5 AND NOT bRamp THEN aCalm[k] := aCalm[k] + 0.01; ELSE aCalm[k] := 0.0; END_IF;
    IF aCalm[k] > 120.0 AND NOT bAnyAlarm AND (aContent[k] < 0.05 OR aContent[k] > 0.95) THEN
        dW := (aDuty[k] - uff) * aP[k] * 0.01 / 600.0;
        IF aContent[k] < 0.05 THEN
            aW0[k] := aW0[k] + dW;
        ELSIF fProd > 1.0 THEN
            u := LIMIT(0.5, aA1[k] + dW / fProd, 1.6);
            dW := (u - aA1[k]) * fProd;  aA1[k] := u;
        END_IF;
        aI[k] := aI[k] - dW / aP[k] / aKc[k] * aTi[k];
    END_IF;
END_FOR;
// time-proportioning, 2 s period: element i of n in a zone conducts in its own slice of the period (phase
// [i/n, i/n + duty)) - the zone gets its duty, the phases see the load spread instead of all at once
fPhase := LMOD(fNow_s / 2.0, 1.0);
FOR j := 0 TO 2 DO aExp[j] := SEL(bRunEnable, 0.0, aFanA[j]); END_FOR;
FOR i := 0 TO 8 DO
    aOn[i] := F_InSlice(fPhase, aElSlice[i], aDuty[aElZone[i]]) AND bRunEnable AND NOT aBroken[i]
              AND aProbe[aElPh[i]] <> i;                       // a probed candidate is held off
    IF aOn[i] THEN aExp[aElPh[i]] := aExp[aElPh[i]] + aElW[i] / 230.0; END_IF;
END_FOR;
GVL_IO.qE1T1 := aOn[0];   // Z1
GVL_IO.qE1T2 := aOn[1];   // Z1
GVL_IO.qE1T3 := aOn[2];   // Z1
GVL_IO.qE1B1 := aOn[3];   // Z1
GVL_IO.qE1B2 := aOn[4];   // Z1
GVL_IO.qE2T1 := aOn[5];   // Z2
GVL_IO.qE2B1 := aOn[6];   // Z2
GVL_IO.qE3T1 := aOn[7];   // Z3
GVL_IO.qE3B1 := aOn[8];   // Z3
GVL_IO.qQF1 := bRunEnable;   // Z1 circulation fan
GVL_IO.qQF2 := bRunEnable;   // Z2 circulation fan
GVL_IO.qQF3 := bRunEnable;   // Z3 circulation fan
// heater break: expected vs measured phase current (oven_ctrl._HeaterBreak, line for line)
FOR i := 0 TO 8 DO
    IF aOn[i] THEN aOnT[i] := fNow_s; END_IF;
    aRecent[i] := fNow_s - aOnT[i] <= 0.3;      // the reading lags: on at some time in t_resp
END_FOR;
FOR j := 0 TO 2 DO
    bSame := TRUE;                                            // same elements on as last cycle?
    FOR i := 0 TO 8 DO IF aElPh[i] = j AND aOn[i] <> aOnLast[i] THEN bSame := FALSE; END_IF; END_FOR;
    IF NOT bSame THEN aSince[j] := fNow_s; END_IF;
    bSettled := ABS(aExp[j] - aExpLag[j]) < 0.1 * aThrA[j];
    aExpLag[j] := aExpLag[j] + (aExp[j] - aExpLag[j]) * 0.01 / 0.100;
    IF aProbe[j] >= 0 THEN                                     // active probe: candidate aProbe[j] held off
        IF fNow_s - aProbeT[j] >= 0.3 THEN aProbeMax[j] := MAX(aProbeMax[j], aExpLag[j] - aMeas[j]); END_IF;
        IF fNow_s - aProbeT[j] >= 2.3 THEN     // a full period: its slice came
            IF aProbeMax[j] < 0.5 * aThrA[j] THEN                  // the short vanished: it is the one
                FOR i := 0 TO 8 DO aCand[i] := aCand[i] AND (aElPh[i] <> j OR i = aProbe[j]); END_FOR;
            ELSE
                aCand[aProbe[j]] := FALSE;
            END_IF;
            aProbe[j] := -1;
        END_IF;
    ELSIF aExpLag[j] - aMeas[j] > aThrA[j] AND fNow_s - aNamedT[j] >= 1.0 THEN   // not while the lagged reading settles after a naming
        aShort[j] := aShort[j] + 0.01;
        FOR i := 0 TO 8 DO
            IF aElPh[i] = j THEN aTry[i] := SEL(aShortOn[j], aRecent[i], aTry[i] AND aRecent[i]) AND NOT aBroken[i]; END_IF;
        END_FOR;
        aShortOn[j] := TRUE;
        IF aShort[j] >= 0.2 THEN
            IF NOT aPhAlarm[j] THEN
                aPhAlarm[j] := TRUE;  aAlarmT[j] := fNow_s;
                FOR i := 0 TO 8 DO IF aElPh[i] = j THEN aCand[i] := aTry[i]; END_IF; END_FOR;
            ELSE
                FOR i := 0 TO 8 DO IF aElPh[i] = j THEN aCand[i] := aCand[i] AND aTry[i]; END_IF; END_FOR;
            END_IF;
        END_IF;
    ELSE
        IF bSettled AND fNow_s - aSince[j] >= 0.3 AND aExpLag[j] - aMeas[j] < 0.2 * aThrA[j] AND aPhAlarm[j] THEN
            FOR i := 0 TO 8 DO
                IF aElPh[i] = j AND aOn[i] THEN aCand[i] := FALSE; END_IF;     // conducted, phase read right: not it
            END_FOR;
        END_IF;
        IF aShort[j] < 0.2 THEN aShortOn[j] := FALSE; END_IF;
        aShort[j] := 0.0;
    END_IF;
    IF aPhAlarm[j] THEN
        n := 0;  m := -1;
        FOR i := 0 TO 8 DO IF aElPh[i] = j AND aCand[i] THEN n := n + 1; IF m < 0 THEN m := i; END_IF; END_IF; END_FOR;
        IF n = 0 THEN                                          // contradiction: start the diagnosis again
            aPhAlarm[j] := FALSE;  aShortOn[j] := FALSE;  aProbe[j] := -1;
        ELSIF n = 1 THEN                                       // named
            IF NOT aBroken[m] THEN aLost[aElZone[m]] := aLost[aElZone[m]] + aElW[m]; END_IF;   // once per element (idempotent)
            aNamedT[j] := fNow_s;
            aBroken[m] := TRUE;  aCand[m] := FALSE;
            aElementAlarm[aElZone[m]] := TRUE;  aPhAlarm[j] := FALSE;  aShortOn[j] := FALSE;  aProbe[j] := -1;
        ELSIF aProbe[j] < 0 AND fNow_s - aAlarmT[j] >= 4.0 THEN
            aProbe[j] := m;  aProbeT[j] := fNow_s;  aProbeMax[j] := -1.0E9;   // the slices cannot tell: probe
        END_IF;
    END_IF;
END_FOR;
FOR i := 0 TO 8 DO aOnLast[i] := aOn[i]; END_FOR;
// a zone whose remaining elements cannot carry the full band at 95% duty: hold the depositor
bHold := FALSE;
FOR k := 0 TO 2 DO
    IF (aP[k] - aLost[k]) * 0.95 < aLoadFull[k] + aW0[k] + (aA1[k] - 1.0) * (aLoadFull[k] - aLoadEmpty[k]) THEN bHold := TRUE; END_IF;
END_FOR;
fPower_W := 0.0;
FOR k := 0 TO 2 DO fPower_W := fPower_W + aDuty[k] * (aP[k] - aLost[k]); END_FOR;
tStable(IN := ABS(aTemp[0] - aSet[0]) < 2.0 AND ABS(aTemp[1] - aSet[1]) < 2.0 AND ABS(aTemp[2] - aSet[2]) < 2.0, PT := T#60S);
bReady := tStable.Q AND NOT bHold;

(* ---- FB_Policy.st ---- *)
// FB_Policy - a learned model evaluated IN the real-time task (TwinCAT 3 Machine Learning inference,
// ONNX, Tc3_MLL FB_MllPrediction - licence TF3800/TF3810 to confirm). Used for fast, bounded decisions:
// drop lead per tube, kick / pass, grip retry. Its output ALWAYS passes FB_SafeEnvelope.
FUNCTION_BLOCK FB_Policy
VAR fbPredict : FB_MllPrediction; END_VAR

(* ---- FB_QC.st ---- *)
// FB_QC - camera verdict (edge PC via ADS: stQc, one per puck) + colour sensor; kick on the fly.
// Camera -> kicker = 110 mm = 5.5 s >= AI latency 0.5 s.
// A rejected cookie is kicked when its puck reaches the kicker (200 ms pulse). Whether it left is
// known at the transfer (I1): until then the puck is 'kicked' and keeps its data.
FUNCTION_BLOCK FB_QC
VAR_IN_OUT aPuck : T_PuckArray; END_VAR
VAR_INPUT fMaster : LREAL; stQc : ST_QcResult; END_VAR
VAR_OUTPUT bKick : BOOL; nKicks, nVerdicts : DINT; END_VAR
VAR fbKick : FB_Arrivals; nSeen, pk : INT; fKickEnd : LREAL; bFirst : BOOL := TRUE; END_VAR
IF bFirst THEN nSeen := stQc.nSeq;  bFirst := FALSE; END_IF;
IF stQc.nSeq <> nSeen THEN                 // a new verdict: 1 pass, 2 reject
    nSeen := stQc.nSeq;  aPuck[stQc.nPuck].nVerdict := stQc.nVerdict;  nVerdicts := nVerdicts + 1;
END_IF;
fbKick(fMaster := fMaster, fStation := 2181.718530718);
IF fbKick.bArrive THEN
    pk := fbKick.nPuck;
    IF aPuck[pk].bFull AND NOT aPuck[pk].bKicked AND aPuck[pk].nVerdict = 2 THEN
        aPuck[pk].bKicked := TRUE;  fKickEnd := fbKick.fArr + 4.0000;  nKicks := nKicks + 1;
    END_IF;
END_IF;
bKick := fMaster < fKickEnd;

(* ---- FB_SafetyIf.st ---- *)
// FB_SafetyIf - the STANDARD side of the TwinSAFE project (EL6910). It never switches a safe
// output: it sends REQUESTS (unlock a door, mute a port, reset) and reads STATUS via the EL6910's
// standard process data. The safety functions themselves (SF1..SF6, SAFETY_CONCEPT.md, safety.py) are
// configured in the TwinSAFE editor from safety/safety_functions.csv.
//   SS1: on any stop demand the NC ramps every axis down (MC_Stop), then TwinSAFE drops K1/K2 after
//        1.20 s (longest ramp + 0.2 s margin, proven in safety.py).
//   Doors S20, S21, S22: unlock request -> TwinSAFE unlocks only after every encoder reports standstill for
//        2.5 s (the standard encoders are a plausibility input; see SAFETY_CONCEPT open items).
//   Ports: airlocks (S-1b) - FB_Airlock sequences them; TwinSAFE enforces the interlocks
//        (outer door unlocks only with the inner side shut and the zone at safe standstill).
FUNCTION_BLOCK FB_SafetyIf
VAR_OUTPUT
    bRunEnable   : BOOL;          // no stop demand active, all doors locked, all resets done
    bStopDemand  : BOOL;          // SS1 in progress -> every station: MC_Stop now
    aDoorLocked  : ARRAY[0..2] OF BOOL;
    aPortMuted   : ARRAY[0..1] OF BOOL;
END_VAR
VAR
    aUnlockReq   : ARRAY[0..2] OF BOOL;   // from the HMI
    aMuteReq     : ARRAY[0..1] OF BOOL;   // from FB_AmrPorts when an AMR is due
END_VAR
bRunEnable := GVL_IO.xSafeRunPermit;      // the EL6910 says: no stop demand, doors locked, resets done
bStopDemand := NOT GVL_IO.xSafeRunPermit;

(* ---- FB_Transfer.st ---- *)
// FB_Transfer - delta C takes the cookies of the row in the pick window (70 mm = 31 s,
// >= 6 takts) in row order (W R B W R B) and places each into the next empty puck on the bend
// (-30..-2 deg). I1 = puck already full (recirculating): skip it, the cookie waits.
// Rows come from FB_Band (the rows really cut); a row is in the window from 1335 mm of band after its cut for
// 70 mm, then it falls off the nose (lost). The band is judged where it was when the puck arrived.
// The grip is known from the vacuum after T_GRAB (0.8 s): held -> the puck is loaded; not held -> the
// cookie stays on the band for the next puck.
FUNCTION_BLOCK FB_Transfer
VAR_IN_OUT stJob : ST_DeltaJob; aPuck : T_PuckArray; END_VAR
VAR_INPUT fMaster : LREAL; fBand : LREAL; nRows : UDINT; fRowPos : LREAL; bPuckFull : BOOL; nVacuum : INT;
    bLoad : BOOL; END_VAR
VAR_OUTPUT bVacuum : BOOL; nLoaded, nGripFail, nRecirc, nEmpty, nLost, nTrackErr : DINT; END_VAR
VAR fbArr : FB_Arrivals; aRow : ARRAY[0..31] OF LREAL; nHead, nTail, nCol, pk, nJobPuck : INT; nSeen : UDINT;
    bFirst : BOOL := TRUE; bWait : BOOL; fGrip, fPlace, d : LREAL;
    aColFlav : ARRAY[0..5] OF INT := [0, 1, 2, 0, 1, 2];   // flavour of each column
END_VAR
IF bFirst THEN nSeen := nRows;  bFirst := FALSE; END_IF;
IF nRows <> nSeen THEN aRow[nTail] := fRowPos;  nTail := (nTail + 1) MOD 32;  nSeen := nRows; END_IF;
fbArr(fMaster := fMaster, fStation := 1550.008729295);
IF bWait AND fMaster >= fGrip THEN         // the grip of the last job
    bWait := FALSE;
    IF nVacuum <= -300 THEN
        aPuck[nJobPuck].bFull := TRUE;  aPuck[nJobPuck].nFlav := aColFlav[nCol];  aPuck[nJobPuck].nCol := nCol;
        aPuck[nJobPuck].fRowPos := aRow[nHead];  aPuck[nJobPuck].nVerdict := 0;
        aPuck[nJobPuck].bKicked := FALSE;  aPuck[nJobPuck].bPending := FALSE;
        nLoaded := nLoaded + 1;  nCol := nCol + 1;
        IF nCol >= 6 THEN nCol := 0;  nHead := (nHead + 1) MOD 32; END_IF;
    ELSE
        nGripFail := nGripFail + 1;  fPlace := fMaster;      // nothing held: vacuum off, the cookie stays
    END_IF;
END_IF;
IF fbArr.bArrive AND bLoad THEN
    pk := fbArr.nPuck;
    d := fBand - (fMaster - fbArr.fArr) * 0.114583333333;   // the band when the puck arrived
    WHILE nHead <> nTail AND d - aRow[nHead] >= 1405.000000000 DO   // past the nose: lost
        nLost := nLost + 6 - INT_TO_DINT(nCol);  nCol := 0;  nHead := (nHead + 1) MOD 32;
    END_WHILE;
    IF bPuckFull THEN                      // recirculating (or a kick that failed: the cookie is still in it)
        nRecirc := nRecirc + 1;
        IF NOT aPuck[pk].bFull THEN nTrackErr := nTrackErr + 1; END_IF;
        aPuck[pk].bKicked := FALSE;
    ELSE
        IF aPuck[pk].bFull AND NOT aPuck[pk].bKicked THEN nTrackErr := nTrackErr + 1; END_IF;
        aPuck[pk].bFull := FALSE;  aPuck[pk].bKicked := FALSE;     // kicked out: empty
        IF nHead = nTail THEN
            nEmpty := nEmpty + 1;
        ELSIF d - aRow[nHead] < 1335.000000000 THEN
            nEmpty := nEmpty + 1;                                     // the next row is not in the window yet
        ELSE
            stJob.nPuck := pk;  stJob.nCol := nCol;  stJob.nLane := -1;  stJob.fRowPos := aRow[nHead];
            stJob.fStart := fbArr.fArr;  stJob.nJob := (stJob.nJob + 1) MOD 10000;
            bWait := TRUE;  nJobPuck := pk;
            fGrip := fbArr.fArr + 16.0000;  fPlace := fbArr.fArr + 40.0000;
        END_IF;
    END_IF;
END_IF;
bVacuum := fMaster < fPlace;

(* ---- MAIN.st ---- *)
// MAIN - one cycle of every station agent; all stations run on ONE time base (the master axis)
PROGRAM MAIN
VAR
    fbMaster  : FB_MasterAxis;
    fbOven    : FB_Oven;          // zones, elements, fans, warm-up gate (oven.py recipe)
    fbBand    : FB_Band;          // band + depositor + topping, geared to the master
    fbTransfer: FB_Transfer;      // delta C: band row -> passing puck, NFC write
    fbQC      : FB_QC;
    fbPickA, fbPickB : FB_DeltaPicker;
    fbLane    : ARRAY[0..2] OF FB_Lane;
    fbPorts   : FB_AmrPorts;
    fbSafety  : FB_SafetyIf;      // S-1: standard side of the TwinSAFE project (requests + status only)
    aPuck     : T_PuckArray;      // what the PLC knows of every puck (filled, flavour, verdict ...)
    aLane     : T_LaneArray;      // per lane: blocked while it indexes, packs to index
END_VAR
fbSafety();                      // first: every station below runs only while fbSafety.bRunEnable
fbMaster(axDrive := GVL_IO.axQ1, axMaster := GVL_IO.axMasterEnc, nEncoder := GVL_IO.encB1);
fbOven(bRunEnable := fbSafety.bRunEnable, aContent := fbBand.aZoneContent);   // last cycle's content
fbBand(axBand := GVL_IO.axQ40, axRolls := GVL_IO.axQ41, axMaster := GVL_IO.axMasterEnc,
       bOvenReady := fbOven.bReady, nDoughLevel := GVL_IO.iolIOL1);
// the stations in the order of the loop: at one master position the transfer comes first, then QC, the kicker,
// delta A, delta B (A and B see their pucks at the same phase: A first)
fbTransfer(stJob := GVL_IO.stDeltaC, aPuck := aPuck, fMaster := fbMaster.fAbs, fBand := fbBand.fPos,
           nRows := fbBand.nRows, fRowPos := fbBand.fRowPos, bPuckFull := GVL_IO.iI1,
           nVacuum := GVL_IO.ioldelta_C_VAC_P, bLoad := GVL_IO.xHmiLoad);
GVL_IO.qdelta_C_VAC := fbTransfer.bVacuum;
fbQC(aPuck := aPuck, fMaster := fbMaster.fAbs, stQc := GVL_IO.stQc);
GVL_IO.qQ18 := fbQC.bKick;
fbPickA(stJob := GVL_IO.stDeltaA, aPuck := aPuck, aLane := aLane, fMaster := fbMaster.fAbs, nDelta := 0,
        fIn := 2534.116936495, fOut := 2629.320124941, nVacuum := GVL_IO.ioldelta_A_VAC_P);
GVL_IO.qdelta_A_VAC := fbPickA.bVacuum;
fbPickB(stJob := GVL_IO.stDeltaB, aPuck := aPuck, aLane := aLane, fMaster := fbMaster.fAbs, nDelta := 1,
        fIn := 2854.116936495, fOut := 2949.320124941, nVacuum := GVL_IO.ioldelta_B_VAC_P);
GVL_IO.qdelta_B_VAC := fbPickB.bVacuum;
fbLane[0](axLane := GVL_IO.axQ20, stLane := aLane[0], fMaster := fbMaster.fAbs);
fbLane[1](axLane := GVL_IO.axQ21, stLane := aLane[1], fMaster := fbMaster.fAbs);
fbLane[2](axLane := GVL_IO.axQ22, stLane := aLane[2], fMaster := fbMaster.fAbs);
fbPorts();
